// TIA Portal V21 export
VAR_GLOBAL   // PLC tag table "Tags_1200"
   BeltStart AT %I0.0 : Bool;   // Belt start button, onboard DI
   BeltStop AT %I0.1 : Bool;   // Belt stop button, onboard DI
   BeltSpeedRaw AT %IW64 : Int;   // Belt speed raw value, onboard AI 0 (0..27648)
   BeltMotor AT %Q0.0 : Bool;   // Belt motor contactor, onboard DQ
END_VAR
